Fanuc KAREL source: KT00137.KL

PROGRAM KT00137
%NOLOCKGROUP
VAR
  R1: REAL
  I2: INTEGER
  OUT: INTEGER
BEGIN
  R1 = 2.0
    I2 = 3
  OUT = R1 DIV I2
END KT00137
